(* IEC 61131-3 sources: PLC_I/plc/src/application, 8 files *)

(* ---- 结构体_运行时.st ---- *)
(* Volatile exchange. Call Server before installed axis consumers each scan.
   ConsumerMask proves program routing, never physical online or safety status. *)
TYPE 结构体_运行时 :
STRUCT
    ast轴 : ARRAY[0..15] OF 结构体_轴状态;
    aw轴命令 : ARRAY[0..15] OF WORD;
    aw轴序列 : ARRAY[0..15] OF WORD;
    adi轴目标 : ARRAY[0..15] OF DINT;
    audi轴速度 : ARRAY[0..15] OF UDINT;
    audi轴加速度 : ARRAY[0..15] OF UDINT;
    audi轴减速度 : ARRAY[0..15] OF UDINT;
    audi轴停止减速度 : ARRAY[0..15] OF UDINT;
    w轴消费掩码 : WORD;
    ast气缸 : ARRAY[0..53] OF 结构体_气缸状态;
    aw气缸命令 : ARRAY[0..53] OF WORD;
    aw气缸序列 : ARRAY[0..53] OF WORD;
    b手动 : BOOL;
    b运行 : BOOL;
    b暂停 : BOOL;
    bHMI在线 : BOOL;
    b复位中 : BOOL;
    (* 上位机命令 2/3/4 的一扫描事件。服务端在受理的同一扫描置位，
       PRG 在下一扫描消费后清零；与物理按钮沿分开，避免被 R_TRIG 合并。 *)
    b启动脉冲 : BOOL;
    b暂停脉冲 : BOOL;
    b恢复脉冲 : BOOL;
    b硬急停 : BOOL;
    b软急停 : BOOL;
    b待复位 : BOOL := TRUE;
    ui输入点数 : UINT;
    ui输出点数 : UINT;
    aw输入 : ARRAY[0..7] OF WORD;
    aw输出 : ARRAY[0..7] OF WORD;
END_STRUCT
END_TYPE

(* ---- 全局变量_错误码.gvl.st ---- *)
(* 拒绝/错误码集中定义。FB 只引用名称，避免数字散落各文件。
   数值与协议 register-map 的拒绝码一致，新增码必须同步协议表。 *)
VAR_GLOBAL CONSTANT
    ERR_已受理   : WORD := 0;
    ERR_签名     : WORD := 1;
    ERR_通信离线 : WORD := 2;
    ERR_急停     : WORD := 3;
    ERR_未绑定   : WORD := 4;
    ERR_离线     : WORD := 5;
    ERR_未使能   : WORD := 6;
    ERR_模式     : WORD := 7;
    ERR_复位中   : WORD := 8;
    ERR_参数     : WORD := 9;
    ERR_忙       : WORD := 10;
    ERR_待复位   : WORD := 11;
    ERR_正式流程 : WORD := 12;
    ERR_未接入   : WORD := 14;
    ERR_非法     : WORD := 15;
    ERR_纪元     : WORD := 16;
    ERR_故障     : WORD := 17;
    ERR_无点位   : WORD := 18;
    ERR_取消     : WORD := 19;
    ERR_定标     : WORD := 20;
    ERR_软限位   : WORD := 21;
    ERR_速度     : WORD := 22;
    ERR_P0       : WORD := 26;
    ERR_目标越限 : WORD := 27;
    ERR_速度无效 : WORD := 28;
END_VAR

(* ---- 函数_动作许可.st ---- *)
(* Sole action-permission boundary (SBR_动作许可 role). Structural validation
   belongs to 函数_校验, never duplicate movement predicates in HMI. *)
FUNCTION 函数_动作许可 : WORD
VAR_INPUT
    Code : WORD;
    ObjectWord : WORD;
    HmiOnline : BOOL;
    JogBusy : BOOL;
    Resetting : BOOL;
    b自动请求 : BOOL := FALSE;
    b气缸已受理 : BOOL := FALSE; (* 仅驱动消费时复核当前许可 *)
    b暂停恢复 : BOOL := FALSE; (* 仅暂停恢复FB的轴27，允许在暂停状态回快照 *)
    b恢复已下发 : BOOL := FALSE; (* 持续复核时忽略本动作自身的Busy *)
    di恢复目标 : DINT := 0;
END_VAR
VAR_IN_OUT
    Runtime : 结构体_运行时;
    Store : 结构体_配置;
END_VAR
VAR
    w类别 : WORD;
    ui对象索引 : UINT;
    ui轴号 : UINT;
    w归属 : WORD;
    b空闲槽 : BOOL;
    b对象已绑定 : BOOL;
    b硬件已接入 : BOOL;
    b是停止 : BOOL;
    b有点位 : BOOL;
    i循环 : UINT;
    i子循环 : UINT;
    di正限位 : DINT;
    di负限位 : DINT;
    di位置 : DINT;
    dw值 : DWORD;
END_VAR

函数_动作许可 := ERR_已受理;
w类别 := SHR(ObjectWord, 8);
ui对象索引 := WORD_TO_UINT(ObjectWord AND 16#00FF);
IF (w类别 > 3) OR ((w类别 = 0) AND (ui对象索引 <> 0))
OR ((w类别 = 1) AND (ui对象索引 >= 16))
OR ((w类别 = 2) AND (ui对象索引 >= 54))
OR ((w类别 = 3) AND (ui对象索引 >= 120)) THEN
    函数_动作许可 := ERR_非法; RETURN;
END_IF;
IF b暂停恢复 AND ((w类别 <> 1) OR (Code <> 27)) THEN
    函数_动作许可 := ERR_非法; RETURN;
END_IF;
ui轴号 := ui对象索引;
b空闲槽 := FALSE;
IF w类别 = 3 THEN
    b空闲槽 := Store.aw点位[ui对象索引, 4] = XJV1_POINT_FREE;
    w归属 := SHR(Store.aw点位[ui对象索引, 4], 2) AND WORD#16#000F;
    ui轴号 := WORD_TO_UINT(w归属);
END_IF;
b对象已绑定 := w类别 = 0;
b硬件已接入 := (Runtime.w轴消费掩码 AND w已绑定轴) = w已绑定轴;
IF w类别 = 1 THEN
    b对象已绑定 := (w已绑定轴 AND SHL(WORD#1, ui轴号)) <> 0;
    b硬件已接入 := (Runtime.w轴消费掩码 AND SHL(WORD#1, ui轴号)) <> 0;
ELSIF w类别 = 3 THEN
    (* An owned point is bound exactly when its owner axis is bound; free
       slots are handled separately below. *)
    b对象已绑定 := NOT b空闲槽 AND ((w已绑定轴 AND SHL(WORD#1, ui轴号)) <> 0);
    b硬件已接入 := (Runtime.w轴消费掩码 AND SHL(WORD#1, ui轴号)) <> 0;
ELSIF w类别 = 2 THEN
    b对象已绑定 := (lw已绑定气缸 AND SHL(LWORD#1, ui对象索引)) <> 0;
    b硬件已接入 := ab气缸映射有效[ui对象索引];
END_IF;
b是停止 := (Code = 9) OR (Code = 10) OR (Code = 26) OR (Code = 42);
(* Stop codes bypass every ordinary gate; an unbound object still rejects 4. *)
IF b是停止 THEN
    IF NOT b对象已绑定 THEN 函数_动作许可 := ERR_未绑定; END_IF;
    RETURN;
END_IF;
IF NOT HmiOnline THEN 函数_动作许可 := ERR_通信离线; RETURN; END_IF;
IF (w类别 = 3) AND b空闲槽 THEN
    (* Free pool slot: only a code-50 claim may address it; the candidate
       owner axis is validated against the binding table in Config. *)
    IF Code <> 50 THEN 函数_动作许可 := ERR_未绑定; RETURN; END_IF;
    IF Runtime.b硬急停 OR Runtime.b软急停 THEN 函数_动作许可 := ERR_急停; RETURN; END_IF;
    IF Resetting THEN 函数_动作许可 := ERR_复位中; RETURN; END_IF;
    IF NOT Runtime.b手动 THEN 函数_动作许可 := ERR_模式; RETURN; END_IF;
    RETURN;
END_IF;
IF Code = 53 THEN 函数_动作许可 := ERR_未接入; RETURN; END_IF;
IF Code = 11 THEN
    (* Clear only the software latch. This does not grant motion permission,
       reset faults, enable an axis, or resume the sequence. *)
    IF Runtime.b硬急停 THEN 函数_动作许可 := ERR_急停; END_IF;
    RETURN;
END_IF;
IF Runtime.b硬急停 OR Runtime.b软急停 THEN 函数_动作许可 := ERR_急停; RETURN; END_IF;
IF NOT b对象已绑定 THEN 函数_动作许可 := ERR_未绑定; RETURN; END_IF;
IF w类别 = 2 THEN
    IF Resetting THEN 函数_动作许可 := ERR_复位中; RETURN; END_IF;
    IF Runtime.b暂停 THEN 函数_动作许可 := ERR_模式; RETURN; END_IF;
    IF b自动请求 THEN
        IF NOT 全局变量_运行配置.b正式流程已接入 THEN 函数_动作许可 := ERR_正式流程; RETURN; END_IF;
        IF NOT Runtime.b运行 THEN 函数_动作许可 := ERR_模式; RETURN; END_IF;
    ELSIF NOT Runtime.b手动 THEN 函数_动作许可 := ERR_模式; RETURN;
    END_IF;
    IF (Code <> 40) AND (Code <> 41) AND (Code <> 50) THEN 函数_动作许可 := ERR_未接入; RETURN; END_IF;
    IF NOT b气缸已受理 AND (全局变量_气缸请求.ast请求[ui对象索引].b忙
        OR Runtime.ast气缸[ui对象索引].b运动中) THEN 函数_动作许可 := ERR_忙; RETURN; END_IF;
    IF Code = 50 THEN RETURN; END_IF;
    IF NOT b硬件已接入 THEN 函数_动作许可 := ERR_未接入; RETURN; END_IF;
    IF NOT ab气缸模块就绪[ui对象索引] THEN 函数_动作许可 := ERR_离线; RETURN; END_IF;
    IF Runtime.ast气缸[ui对象索引].b故障 THEN 函数_动作许可 := ERR_故障; RETURN; END_IF;
    (* 手动调试不依赖上电复位和现场配置确认：手动模式下可以直接触发
       动点/原点。自动请求仍必须完成确认与复位，避免工艺在未确认配置上运行。 *)
    IF b自动请求 THEN
        IF Runtime.b待复位 THEN 函数_动作许可 := ERR_待复位; RETURN; END_IF;
        IF NOT Store.b已确认 THEN 函数_动作许可 := ERR_未接入; RETURN; END_IF;
    END_IF;
    IF NOT 气缸_配置有效(缸号 := ui对象索引, Store := Store) THEN 函数_动作许可 := ERR_参数; END_IF;
    RETURN;
END_IF;
(* 整机启动/暂停/恢复。正式工艺未接入时三条一律拒绝 12，与原程序
   “NOT b正式流程已接入 → 拒绝” 一致；接入后由运行状态机判定模式与暂停，
   这里只做安全与前置条件检查，不复制运行状态机的优先级逻辑。 *)
IF (Code = 2) OR (Code = 3) OR (Code = 4) THEN
    IF NOT 全局变量_运行配置.b正式流程已接入 THEN 函数_动作许可 := ERR_正式流程; RETURN; END_IF;
    IF Code = 2 THEN
        IF Runtime.b待复位 THEN 函数_动作许可 := ERR_未接入; RETURN; END_IF;
    ELSIF Code = 4 THEN
        IF NOT Runtime.b暂停 THEN 函数_动作许可 := ERR_未接入; RETURN; END_IF;
    END_IF;
    RETURN;
END_IF;
IF Resetting AND (Code <> 21) THEN 函数_动作许可 := ERR_复位中; RETURN; END_IF;
IF w类别 = 0 THEN
    IF Code = 1 THEN
        IF NOT b硬件已接入 THEN 函数_动作许可 := ERR_未接入; RETURN; END_IF;
        FOR i循环 := 0 TO 15 DO
            IF (w已绑定轴 AND SHL(WORD#1, i循环)) <> 0 THEN
                IF NOT Runtime.ast轴[i循环].b在线 THEN 函数_动作许可 := ERR_离线; RETURN; END_IF;
            END_IF;
        END_FOR;
    ELSIF Code = 52 THEN
        IF NOT Runtime.b手动 THEN 函数_动作许可 := ERR_模式; RETURN; END_IF;
        FOR i循环 := 0 TO 15 DO
            IF (w已绑定轴 AND SHL(WORD#1, i循环)) <> 0 THEN
                IF NOT Runtime.ast轴[i循环].b在线 THEN 函数_动作许可 := ERR_离线; RETURN; END_IF;
                IF Runtime.ast轴[i循环].b故障 THEN 函数_动作许可 := ERR_故障; RETURN; END_IF;
                IF Runtime.ast轴[i循环].b运动中 OR NOT Runtime.ast轴[i循环].b静止 THEN
                    函数_动作许可 := ERR_忙; RETURN;
                END_IF;
                di正限位 := DWORD_TO_DINT(SHL(WORD_TO_DWORD(Store.aw轴配置[i循环, 0]), 16) OR WORD_TO_DWORD(Store.aw轴配置[i循环, 1]));
                di负限位 := DWORD_TO_DINT(SHL(WORD_TO_DWORD(Store.aw轴配置[i循环, 2]), 16) OR WORD_TO_DWORD(Store.aw轴配置[i循环, 3]));
                IF (Store.aw轴配置[i循环, 14] <> 1) OR (Store.aw轴配置[i循环, 15] <> 0) THEN
                    函数_动作许可 := ERR_定标; RETURN;
                END_IF;
                IF di负限位 >= di正限位 THEN 函数_动作许可 := ERR_软限位; RETURN; END_IF;
                FOR i子循环 := 2 TO 6 DO
                    dw值 := SHL(WORD_TO_DWORD(Store.aw轴配置[i循环, i子循环 * 2]), 16) OR WORD_TO_DWORD(Store.aw轴配置[i循环, i子循环 * 2 + 1]);
                    IF (dw值 = 0) OR (dw值 > DWORD#2147483647) THEN
                        函数_动作许可 := 函数_参数码(i子循环); RETURN;
                    END_IF;
                    IF NOT 函数_额定值(AxisIndex := i循环, Field := i子循环,
                        Value := DWORD_TO_UDINT(dw值)) THEN
                        函数_动作许可 := 函数_参数码(i子循环); RETURN;
                    END_IF;
                END_FOR;
                (* Standby point P0 of axis i is pool slot i by definition. *)
                IF (SHR(Store.aw点位[i循环, 4], 2) AND WORD#16#000F) <> UINT_TO_WORD(i循环)
                OR (Store.aw点位[i循环, 4] AND 3) <> 3 THEN 函数_动作许可 := ERR_无点位; RETURN; END_IF;
                di位置 := DWORD_TO_DINT(SHL(WORD_TO_DWORD(Store.aw点位[i循环, 0]), 16) OR WORD_TO_DWORD(Store.aw点位[i循环, 1]));
                dw值 := SHL(WORD_TO_DWORD(Store.aw点位[i循环, 2]), 16) OR WORD_TO_DWORD(Store.aw点位[i循环, 3]);
                IF (di位置 < di负限位) OR (di位置 > di正限位) THEN 函数_动作许可 := ERR_P0; RETURN; END_IF;
                IF (dw值 = 0) OR (dw值 > DWORD#2147483647) THEN 函数_动作许可 := ERR_速度无效; RETURN; END_IF;
            END_IF;
        END_FOR;
        FOR i循环 := 0 TO 53 DO
            IF (lw已绑定气缸 AND SHL(LWORD#1, i循环)) <> 0 THEN
                IF NOT 气缸_配置有效(缸号 := i循环, Store := Store) THEN 函数_动作许可 := ERR_参数; RETURN; END_IF;
                IF 全局变量_气缸请求.ast请求[i循环].b忙 THEN 函数_动作许可 := ERR_忙; RETURN; END_IF;
            END_IF;
        END_FOR;
    ELSE
        函数_动作许可 := ERR_未接入;
    END_IF;
    RETURN;
END_IF;
IF (Runtime.aw轴命令[ui轴号] <> 0) AND (Code <> 21) THEN
    函数_动作许可 := ERR_忙; RETURN;
END_IF;
IF NOT b自动请求 AND 全局变量_轴请求.ast请求[ui轴号].b忙 AND (Code <> 21) THEN
    函数_动作许可 := ERR_忙; RETURN;
END_IF;
CASE Code OF
    20, 21, 22, 23, 24, 25, 27, 28, 29, 30, 31, 50: ;
ELSE
    函数_动作许可 := ERR_未接入; RETURN;
END_CASE;
IF NOT Runtime.ast轴[ui轴号].b在线 THEN 函数_动作许可 := ERR_离线; RETURN; END_IF;
(* 硬限位未接线时必须保留软限位，否则拒绝运动类命令，避免无边界保护。 *)
IF (Code = 22) OR (Code = 24) OR (Code = 25) OR (Code = 27)
    OR (Code = 28) OR (Code = 29) THEN
    IF NOT 全局变量_运行配置.b硬限位已接线
        AND ((Store.aw轴配置[ui轴号, 14] AND WORD#16#0001) = 0) THEN
        函数_动作许可 := ERR_未接入; RETURN;
    END_IF;
END_IF;
(* 写参数（31/50）不动轴，报警期间也允许改；复位 23 与去使能 21 同样放行。 *)
IF Runtime.ast轴[ui轴号].b故障 AND (Code <> 21) AND (Code <> 23)
    AND (Code <> 31) AND (Code <> 50) THEN
    函数_动作许可 := ERR_故障; RETURN;
END_IF;
IF b暂停恢复 THEN
    (* 恢复有独立模式条件；不能借普通自动许可放开暂停中的其他命令。 *)
    IF NOT 全局变量_运行配置.b正式流程已接入 THEN 函数_动作许可 := ERR_正式流程; RETURN; END_IF;
    (* 运行控制在暂停时发布手动模式，恢复仍以暂停握手为准。 *)
    IF NOT Runtime.b暂停 THEN 函数_动作许可 := ERR_模式; RETURN; END_IF;
    IF Runtime.b待复位 THEN 函数_动作许可 := ERR_待复位; RETURN; END_IF;
    di正限位 := DWORD_TO_DINT(SHL(WORD_TO_DWORD(Store.aw轴配置[ui轴号, 0]), 16) OR WORD_TO_DWORD(Store.aw轴配置[ui轴号, 1]));
    di负限位 := DWORD_TO_DINT(SHL(WORD_TO_DWORD(Store.aw轴配置[ui轴号, 2]), 16) OR WORD_TO_DWORD(Store.aw轴配置[ui轴号, 3]));
    IF (Store.aw轴配置[ui轴号, 14] AND 1) <> 0 THEN
        IF (di负限位 >= di正限位) OR (di恢复目标 < di负限位) OR (di恢复目标 > di正限位) THEN
            函数_动作许可 := ERR_软限位; RETURN;
        END_IF;
    END_IF;
    IF ((di恢复目标 > Runtime.ast轴[ui轴号].di位置) AND ((Runtime.ast轴[ui轴号].w限位 AND 5) <> 0))
        OR ((di恢复目标 < Runtime.ast轴[ui轴号].di位置) AND ((Runtime.ast轴[ui轴号].w限位 AND 10) <> 0)) THEN
        函数_动作许可 := ERR_故障; RETURN;
    END_IF;
ELSIF b自动请求 THEN
    IF NOT 全局变量_运行配置.b正式流程已接入 THEN 函数_动作许可 := ERR_正式流程; RETURN; END_IF;
    IF NOT Runtime.b运行 OR Runtime.b暂停 THEN 函数_动作许可 := ERR_模式; RETURN; END_IF;
    IF Runtime.b待复位 THEN 函数_动作许可 := ERR_待复位; RETURN; END_IF;
ELSIF NOT Runtime.b手动 AND (Code <> 21) THEN 函数_动作许可 := ERR_模式; RETURN;
END_IF;
IF ((Code = 22) OR (Code = 24) OR (Code = 25) OR (Code = 27) OR (Code = 28) OR (Code = 29) OR (Code = 30))
AND NOT Runtime.ast轴[ui轴号].b已使能 THEN 函数_动作许可 := ERR_未使能; RETURN; END_IF;
(* 清故障在报警态必须可重试：轴停在 ErrorStop 时 b运动中 可能因残留停止阶段为真，
   若因此拒绝 23，现场就永远清不掉。复位本身仍要求 MC_Reset 成功。 *)
IF (Code >= 20) AND (Code <= 30) AND (Code <> 21)
AND NOT (b暂停恢复 AND b恢复已下发)
AND NOT Runtime.ast轴[ui轴号].b可下发 THEN
    函数_动作许可 := ERR_忙; RETURN;
END_IF;
IF (Runtime.ast轴[ui轴号].b运动中 OR NOT Runtime.ast轴[ui轴号].b静止) AND (Code <> 21) AND (Code <> 23)
    AND NOT (b暂停恢复 AND b恢复已下发) THEN
    函数_动作许可 := ERR_忙; RETURN;
END_IF;
IF (Code = 24) OR (Code = 25) THEN
    IF JogBusy THEN 函数_动作许可 := ERR_忙; RETURN; END_IF;
    IF ((Code = 24) AND ((Runtime.ast轴[ui轴号].w限位 AND 5) <> 0))
    OR ((Code = 25) AND ((Runtime.ast轴[ui轴号].w限位 AND 10) <> 0)) THEN
        函数_动作许可 := ERR_故障; RETURN;
    END_IF;
END_IF;
IF Code = 29 THEN
    b有点位 := FALSE;
    FOR i循环 := 0 TO 119 DO
        b有点位 := b有点位 OR ((SHR(Store.aw点位[i循环, 4], 2) AND WORD#16#000F) = UINT_TO_WORD(ui轴号)
            AND ((Store.aw点位[i循环, 4] AND 3) = 3));
    END_FOR;
    IF NOT b有点位 THEN 函数_动作许可 := ERR_无点位; RETURN; END_IF;
END_IF;
IF ((Code >= 20) AND (Code <= 30)) AND NOT b硬件已接入 THEN
    函数_动作许可 := ERR_未接入; RETURN;
END_IF;
IF (Code = 20) OR (Code = 22) OR (Code = 24) OR (Code = 25)
OR (Code = 27) OR (Code = 28) OR (Code = 29) THEN
    FOR i子循环 := 2 TO 6 DO
        dw值 := SHL(WORD_TO_DWORD(Store.aw轴配置[ui轴号, i子循环 * 2]), 16)
            OR WORD_TO_DWORD(Store.aw轴配置[ui轴号, i子循环 * 2 + 1]);
        IF NOT 函数_额定值(AxisIndex := ui轴号, Field := i子循环,
            Value := DWORD_TO_UDINT(dw值)) THEN
            函数_动作许可 := 函数_参数码(i子循环); RETURN;
        END_IF;
    END_FOR;
END_IF;
END_FUNCTION

(* ---- 功能块_暂停恢复.st ---- *)
(* 暂停快照与恢复。移植自原程序“暂停快照 / 暂停回位”三段，只保留必要行为：

   暂停沿 -> 对运动中轴下受控停止 26 -> 全部静止后抓拍位置
   恢复请求 -> 对偏离超过容差的轴下发绝对定位 27 回快照位置 -> 结果 2 即完成
   急停 / 轴离线或故障 -> 立即判失败并撤销本块下发的命令

   不产生动作许可，不替代 功能块_轴 的安全判定。
   必须在 功能块_服务端 之后、各轴消费之前调用（服务端每扫描开头清零命令数组）。 *)
FUNCTION_BLOCK 功能块_暂停恢复
VAR_INPUT
    b暂停 : BOOL;
    b请求 : BOOL;
    b急停 : BOOL;
    di容差 : DINT;
    (* 停稳确认时间。原程序为 300 ms；做成输入便于自测用更短的值，
       现场调用保持 300 ms。 *)
    di停稳ms : DINT;
END_VAR
VAR_IN_OUT
    Runtime : 结构体_运行时;
END_VAR
VAR_OUTPUT
    b恢复中 : BOOL;
    b恢复完成 : BOOL;
    b恢复失败 : BOOL;
    b曾偏离 : BOOL;
    b已抓拍 : BOOL;
    (* 内部阶段只读发布，供上位机诊断与自测观察。 *)
    ui内部阶段 : UINT;
END_VAR
VAR
    i阶段 : UINT; (* 0 空闲，1 停车等待静止，2 已抓拍待恢复，3 回位中 *)
    b暂停上周期 : BOOL;
    b请求上周期 : BOOL;
    b请求沿 : BOOL;
    adi快照 : ARRAY[0..15] OF DINT;
    (* 只有收到本轮回位 27 的轴才参与完成判定；未偏离的轴不动作，
       不能被当成“未到位”而把恢复永久卡住。 *)
    ab已下发 : ARRAY[0..15] OF BOOL;
    w序列 : WORD;
    b暂停沿 : BOOL;
    b封锁 : BOOL;
    b全部静止 : BOOL;
    b全部到位 : BOOL;
    b取消恢复 : BOOL;
    b恢复动作存在 : BOOL;
    w许可 : WORD;
    tmr停稳 : TON;
    tmr恢复 : TON;
    i循环 : UINT;
END_VAR

b恢复中 := FALSE;
b取消恢复 := (i阶段 = 3) AND (NOT b暂停 OR NOT b请求);
(* b已抓拍 是锁存状态，不是脉冲：暂停沿/解除时清零，抓拍成功时置位。
   上位机与自测都靠它判断“快照是否有效”，脉冲化会漏读。 *)
b暂停沿 := b暂停 AND NOT b暂停上周期;
b暂停上周期 := b暂停;
b请求沿 := b请求 AND NOT b请求上周期;
b请求上周期 := b请求;

(* 安全条件不满足时任何恢复都不成立。 *)
b封锁 := b急停 OR Runtime.b硬急停 OR Runtime.b软急停;
IF b请求沿 OR (i阶段 = 3) THEN
    b封锁 := b封锁 OR NOT Runtime.bHMI在线 OR Runtime.b待复位 OR Runtime.b复位中
        OR NOT 全局变量_运行配置.b正式流程已接入;
END_IF;
FOR i循环 := 0 TO 15 DO
    IF (w已绑定轴 AND SHL(WORD#1, i循环)) <> 0 THEN
        b封锁 := b封锁 OR NOT Runtime.ast轴[i循环].b在线 OR Runtime.ast轴[i循环].b故障;
    END_IF;
END_FOR;
(* 先完整预检全部目标，再发任何轴；回位中每扫描继续复核。
   使用LINT比较，DINT极值两端相减不会溢出。 *)
IF ((i阶段 = 2) AND b请求沿) OR (i阶段 = 3) THEN
    FOR i循环 := 0 TO 15 DO
        IF (w已绑定轴 AND SHL(WORD#1, i循环)) <> 0 THEN
            IF ab已下发[i循环] OR
                (ABS(DINT_TO_LINT(Runtime.ast轴[i循环].di位置) - DINT_TO_LINT(adi快照[i循环])) > DINT_TO_LINT(di容差)) THEN
                w许可 := 函数_动作许可(Code := 27, ObjectWord := WORD#16#0100 OR UINT_TO_WORD(i循环),
                    HmiOnline := Runtime.bHMI在线, JogBusy := FALSE, Resetting := Runtime.b复位中,
                    b暂停恢复 := TRUE, b恢复已下发 := (i阶段 = 3) AND ab已下发[i循环],
                    di恢复目标 := adi快照[i循环], Runtime := Runtime, Store := 全局变量_保持区.Store);
                b封锁 := b封锁 OR (w许可 <> 0);
            END_IF;
        END_IF;
    END_FOR;
END_IF;
IF (i阶段 = 3) AND b封锁 THEN b取消恢复 := TRUE; END_IF;

IF b暂停沿 THEN
    i阶段 := 1;
    b曾偏离 := FALSE;
    b恢复完成 := FALSE;
    b恢复失败 := FALSE;
    b已抓拍 := FALSE;
    w序列 := w序列 + 1;
    tmr停稳(IN := FALSE, PT := DINT_TO_TIME(di停稳ms));
    FOR i循环 := 0 TO 15 DO
        adi快照[i循环] := Runtime.ast轴[i循环].di位置;
        ab已下发[i循环] := FALSE;
    END_FOR;
ELSIF NOT b暂停 THEN
    i阶段 := 0;
    b曾偏离 := FALSE;
    b已抓拍 := FALSE;
END_IF;

CASE i阶段 OF
    1:
        (* 受控停止。序列固定，重复下发同一序列不会在轴内重复触发。 *)
        b全部静止 := TRUE;
        FOR i循环 := 0 TO 15 DO
            IF (w已绑定轴 AND SHL(WORD#1, i循环)) <> 0 THEN
                IF Runtime.ast轴[i循环].b运动中 OR NOT Runtime.ast轴[i循环].b静止 THEN
                    b全部静止 := FALSE;
                    Runtime.aw轴命令[i循环] := 26;
                    Runtime.aw轴序列[i循环] := w序列;
                END_IF;
            END_IF;
        END_FOR;
        tmr停稳(IN := b全部静止 AND NOT b封锁, PT := DINT_TO_TIME(di停稳ms));
        IF tmr停稳.Q THEN
            (* 停稳后重新抓拍：减速距离不算偏离。 *)
            FOR i循环 := 0 TO 15 DO adi快照[i循环] := Runtime.ast轴[i循环].di位置; END_FOR;
            b已抓拍 := TRUE;
            i阶段 := 2;
        END_IF;
    2:
        (* 暂停期间只监视偏离，不自动动作。 *)
        FOR i循环 := 0 TO 15 DO
            IF (w已绑定轴 AND SHL(WORD#1, i循环)) <> 0 THEN
                IF ABS(DINT_TO_LINT(Runtime.ast轴[i循环].di位置) - DINT_TO_LINT(adi快照[i循环])) > DINT_TO_LINT(di容差) THEN
                    b曾偏离 := TRUE;
                END_IF;
            END_IF;
        END_FOR;
        (* 恢复请求只在上升沿处理一次：b请求 是电平，重复处理会每扫描
           重新下发 27，命令槽无法释放，安全封锁时也撤不干净。 *)
        IF b请求沿 AND b封锁 THEN b恢复失败 := TRUE; END_IF;
        IF b请求沿 AND NOT b封锁 THEN
            b恢复完成 := FALSE;
            b恢复失败 := FALSE;
            b恢复动作存在 := FALSE;
            FOR i循环 := 0 TO 15 DO
                IF ((w已绑定轴 AND SHL(WORD#1, i循环)) <> 0)
                    AND (ABS(DINT_TO_LINT(Runtime.ast轴[i循环].di位置) - DINT_TO_LINT(adi快照[i循环])) > DINT_TO_LINT(di容差)) THEN
                    b恢复动作存在 := TRUE;
                END_IF;
            END_FOR;
            IF b恢复动作存在 THEN
                w序列 := w序列 + 1;
                FOR i循环 := 0 TO 15 DO ab已下发[i循环] := FALSE; END_FOR;
                FOR i循环 := 0 TO 15 DO
                    IF (w已绑定轴 AND SHL(WORD#1, i循环)) <> 0 THEN
                        IF ABS(DINT_TO_LINT(Runtime.ast轴[i循环].di位置) - DINT_TO_LINT(adi快照[i循环])) > DINT_TO_LINT(di容差) THEN
                            (* 回位参数取保持配置，与命令 27 的下发参数同源。 *)
                            Runtime.adi轴目标[i循环] := adi快照[i循环];
                            Runtime.audi轴速度[i循环] := DWORD_TO_UDINT(
                                SHL(WORD_TO_DWORD(全局变量_保持区.Store.aw轴配置[i循环, 4]), 16)
                                OR WORD_TO_DWORD(全局变量_保持区.Store.aw轴配置[i循环, 5]));
                            Runtime.audi轴加速度[i循环] := DWORD_TO_UDINT(
                                SHL(WORD_TO_DWORD(全局变量_保持区.Store.aw轴配置[i循环, 8]), 16)
                                OR WORD_TO_DWORD(全局变量_保持区.Store.aw轴配置[i循环, 9]));
                            Runtime.audi轴减速度[i循环] := DWORD_TO_UDINT(
                                SHL(WORD_TO_DWORD(全局变量_保持区.Store.aw轴配置[i循环, 10]), 16)
                                OR WORD_TO_DWORD(全局变量_保持区.Store.aw轴配置[i循环, 11]));
                            Runtime.audi轴停止减速度[i循环] := DWORD_TO_UDINT(
                                SHL(WORD_TO_DWORD(全局变量_保持区.Store.aw轴配置[i循环, 12]), 16)
                                OR WORD_TO_DWORD(全局变量_保持区.Store.aw轴配置[i循环, 13]));
                            Runtime.aw轴命令[i循环] := 27;
                            Runtime.aw轴序列[i循环] := w序列;
                            ab已下发[i循环] := TRUE;
                        END_IF;
                    END_IF;
                END_FOR;
                tmr恢复(IN := FALSE, PT := T#120s);
                i阶段 := 3;
            ELSE
                (* 没偏离就没有要回的位置，恢复直接成立。 *)
                b恢复完成 := TRUE;
            END_IF;
        END_IF;

    3:
        b恢复中 := TRUE;
        b全部到位 := TRUE;
        FOR i循环 := 0 TO 15 DO
            IF (w已绑定轴 AND SHL(WORD#1, i循环)) <> 0 AND ab已下发[i循环] THEN
                b全部到位 := b全部到位 AND (Runtime.ast轴[i循环].w序列 = w序列)
                    AND (Runtime.ast轴[i循环].w运动结果 = 2)
                    AND Runtime.ast轴[i循环].b静止;
            END_IF;
        END_FOR;
        tmr恢复(IN := TRUE, PT := T#120s);
        IF b取消恢复 OR b封锁 OR tmr恢复.Q THEN
            b取消恢复 := TRUE;
            b恢复失败 := TRUE;
            b恢复中 := FALSE;
            i阶段 := 2;
        ELSIF b全部到位 THEN
            FOR i循环 := 0 TO 15 DO ab已下发[i循环] := FALSE; END_FOR;
            b恢复完成 := TRUE;
            b恢复中 := FALSE;
            i阶段 := 2;
        END_IF;
END_CASE;
(* 清命令槽不能取消轴内已锁存的27；主动发26并使用新序列。 *)
IF b取消恢复 THEN
    w序列 := w序列 + 1;
    FOR i循环 := 0 TO 15 DO
        IF ab已下发[i循环] THEN
            Runtime.aw轴命令[i循环] := 26;
            Runtime.aw轴序列[i循环] := w序列;
            ab已下发[i循环] := FALSE;
        END_IF;
    END_FOR;
    b恢复中 := FALSE;
    b恢复完成 := FALSE;
    b恢复失败 := TRUE;
END_IF;
ui内部阶段 := i阶段;
END_FUNCTION_BLOCK

(* ---- 功能块_模式管理.st ---- *)
(* 模式/暂停恢复的唯一状态拥有者。服务端之后、轴组之前调用一次。 *)
FUNCTION_BLOCK 功能块_模式管理
VAR_INPUT StartButton : BOOL; PauseButton : BOOL; ResetButton : BOOL; END_VAR
VAR_IN_OUT Runtime : 结构体_运行时; END_VAR
VAR
    fb运行 : 功能块_运行控制;
    fb暂停恢复 : 功能块_暂停恢复;
    fb启动滤波 : 功能块_输入滤波;
    fb暂停滤波 : 功能块_输入滤波;
    fb复位滤波 : 功能块_输入滤波;
    b复位事件 : BOOL;
    b复位上周期 : BOOL;
    b设备报警 : BOOL;
    b急停 : BOOL;
    i循环 : UINT;
END_VAR
fb启动滤波(b信号 := StartButton, i模式 := 1,
    di滤波时间真 := 全局变量_运行配置.di输入滤波时间ms,
    di滤波时间假 := 全局变量_运行配置.di输入滤波时间ms);
fb暂停滤波(b信号 := PauseButton, i模式 := 1,
    di滤波时间真 := 全局变量_运行配置.di输入滤波时间ms,
    di滤波时间假 := 全局变量_运行配置.di输入滤波时间ms);
fb复位滤波(b信号 := ResetButton, i模式 := 1,
    di滤波时间真 := 全局变量_运行配置.di输入滤波时间ms,
    di滤波时间假 := 全局变量_运行配置.di输入滤波时间ms);
b复位事件 := fb复位滤波.b滤波信号 AND NOT b复位上周期;
b复位上周期 := fb复位滤波.b滤波信号;
b急停 := Runtime.b硬急停;
(* ===== 区域 3：运行模式与命令脉冲消费 ===== *)
(* 运行状态机：物理按钮 + 上位机命令 2/3/4。命令 2 在
   b正式流程已接入 = FALSE 时仍由 函数_动作许可 拒绝为 12。 *)
b设备报警 := FALSE;
FOR i循环 := 0 TO 15 DO
    IF (w已绑定轴 AND SHL(WORD#1, i循环)) <> 0 THEN b设备报警 := b设备报警 OR Runtime.ast轴[i循环].b故障; END_IF;
END_FOR;
fb运行(b初始化完成 := TRUE,
    b系统复位完成 := NOT Runtime.b待复位,
    b系统复位中 := FALSE,
    b系统复位失败 := FALSE,
    b启动按钮 := fb启动滤波.b滤波信号 AND 全局变量_运行配置.b正式流程已接入,
    b暂停按钮 := fb暂停滤波.b滤波信号,
    b启动事件 := Runtime.b启动脉冲,
    b暂停事件 := Runtime.b暂停脉冲,
    (* 物理复位按钮与命令 4 等效：原程序“暂停中按复位进入暂停恢复”。 *)
    b恢复事件 := Runtime.b恢复脉冲 OR (b复位事件 AND 全局变量_运行配置.b正式流程已接入),
    b致命报警 := Runtime.b硬急停 OR Runtime.b软急停 OR b设备报警,
    b急停 := b急停 OR Runtime.b软急停,
    b暂停报警 := b设备报警,
    b预警 := FALSE,
    b暂停恢复中 := fb暂停恢复.b恢复中,
    b暂停恢复完成 := fb暂停恢复.b恢复完成,
    b暂停恢复失败 := fb暂停恢复.b恢复失败,
    b流程完成 := FALSE);
Runtime.b运行 := fb运行.b运行指令;
Runtime.b暂停 := fb运行.b暂停中;
Runtime.b手动 := fb运行.b手动模式;
(* 命令 2/3/4 是一扫描事件：服务端本扫描置位，这里消费后立即清零，
   下一扫描不会重复触发。 *)
Runtime.b启动脉冲 := FALSE;
Runtime.b暂停脉冲 := FALSE;
Runtime.b恢复脉冲 := FALSE;

(* 暂停编排：必须在服务端之后，服务端每扫描开头清零命令数组。 *)
fb暂停恢复(b暂停 := fb运行.b暂停中, b请求 := fb运行.b暂停恢复请求,
    b急停 := b急停,
    di容差 := 全局变量_运行配置.di暂停恢复容差,
    di停稳ms := 全局变量_运行配置.di暂停停稳ms, Runtime := Runtime);

(* Cancel automatic requests before consumers when mode changes in this scan.
   Preserve existing stop/disable/reset pulses from the Server. *)
FOR i循环 := 0 TO 15 DO
    IF 全局变量_轴请求.ast请求[i循环].b忙
    AND 全局变量_轴请求.ast请求[i循环].b已下发
    AND (全局变量_轴请求.ast请求[i循环].w命令 <> 26)
    AND (NOT Runtime.b运行 OR Runtime.b暂停 OR NOT Runtime.bHMI在线
        OR Runtime.b硬急停 OR Runtime.b软急停
        OR Runtime.b待复位 OR Runtime.b复位中) THEN
        IF (Runtime.aw轴命令[i循环] = 0) OR (Runtime.aw轴命令[i循环] = 22)
        OR (Runtime.aw轴命令[i循环] = 27) THEN
            Runtime.aw轴命令[i循环] := 26;
        END_IF;
    END_IF;
END_FOR;

END_FUNCTION_BLOCK

(* ---- 功能块_系统复位.st ---- *)
(* Owns reset phase, committed sequence and timeout. Operation 0 advances once
   before arbitration; 1 accepts reset; 2 cancels immediately during arbitration.
   Start/cancel never advance the timer or phase machine a second time. *)
FUNCTION_BLOCK 功能块_系统复位
VAR_INPUT
    Operation : UINT;
    Sequence : WORD;
END_VAR
VAR_IN_OUT
    Runtime : 结构体_运行时;
END_VAR
VAR_OUTPUT
    Busy : BOOL;
    StopRequested : BOOL;
    Failed : BOOL;
END_VAR
VAR
    ui复位阶段 : UINT;
    w复位序列 : WORD;
    b复位完成 : BOOL;
    b复位失败 : BOOL;
    tmr复位 : TON;
    i循环 : UINT;
END_VAR

StopRequested := FALSE;
Failed := FALSE;
CASE Operation OF
    1:
        Runtime.b待复位 := TRUE;
        w复位序列 := Sequence;
        ui复位阶段 := 1;
        StopRequested := TRUE;
    2:
        ui复位阶段 := 0;
    0:
        tmr复位(IN := ui复位阶段 <> 0, PT := T#30s);
        b复位失败 := Runtime.b硬急停 OR Runtime.b软急停 OR tmr复位.Q;
        FOR i循环 := 0 TO 15 DO
            IF (w已绑定轴 AND SHL(WORD#1, i循环)) <> 0 THEN
                b复位失败 := b复位失败 OR NOT Runtime.ast轴[i循环].b在线;
            END_IF;
        END_FOR;
        IF (ui复位阶段 <> 0) AND b复位失败 THEN
            ui复位阶段 := 0;
            Runtime.b待复位 := TRUE;
            StopRequested := TRUE;
            Failed := TRUE;
        END_IF;
        CASE ui复位阶段 OF
            1:
                b复位完成 := TRUE;
                FOR i循环 := 0 TO 15 DO
                    IF (w已绑定轴 AND SHL(WORD#1, i循环)) <> 0 THEN
                        b复位完成 := b复位完成 AND NOT Runtime.ast轴[i循环].b运动中
                            AND Runtime.ast轴[i循环].b可下发
                            AND (Runtime.ast轴[i循环].b静止 OR (Runtime.ast轴[i循环].b故障 AND (Runtime.ast轴[i循环].di速度 = 0)));
                    END_IF;
                END_FOR;
                IF b复位完成 THEN ui复位阶段 := 2; END_IF;
            2:
                FOR i循环 := 0 TO 15 DO
                    IF (w已绑定轴 AND SHL(WORD#1, i循环)) <> 0 THEN
                        Runtime.aw轴命令[i循环] := 23;
                        Runtime.aw轴序列[i循环] := w复位序列;
                    END_IF;
                END_FOR;
                ui复位阶段 := 3;
            3:
                b复位完成 := TRUE;
                FOR i循环 := 0 TO 15 DO
                    IF (w已绑定轴 AND SHL(WORD#1, i循环)) <> 0 THEN
                        b复位完成 := b复位完成 AND (Runtime.ast轴[i循环].w序列 = w复位序列)
                            AND (Runtime.ast轴[i循环].w运动结果 = 2) AND NOT Runtime.ast轴[i循环].b故障
                            AND Runtime.ast轴[i循环].b静止 AND NOT Runtime.ast轴[i循环].b运动中;
                    END_IF;
                END_FOR;
                IF b复位完成 THEN Runtime.b待复位 := FALSE; ui复位阶段 := 4; END_IF;
            4: ui复位阶段 := 0;
        END_CASE;
END_CASE;
Busy := ui复位阶段 <> 0;
END_FUNCTION_BLOCK

(* ---- 功能块_输入滤波.st ---- *)
(* 现场输入去抖。语义与原程序 功能块_输入滤波 一致：
   模式 0 直通；模式 1 按真/假时间分别计时，先到者生效。
   安全输入（急停 X3）不经过本块，避免滤波延迟安全响应。
   X0/X1/X2 走 20 ms 去抖，与原程序 子程序_IO映射__采集 一致。 *)
FUNCTION_BLOCK 功能块_输入滤波
VAR_INPUT
    b信号 : BOOL;
    i模式 : INT; (* 0 = 直通，1 = 去抖 *)
    di滤波时间真 : DINT; (* ms *)
    di滤波时间假 : DINT; (* ms *)
END_VAR
VAR_OUTPUT
    b滤波信号 : BOOL;
END_VAR
VAR
    tmr延时真 : TON;
    tmr延时假 : TON;
END_VAR

CASE i模式 OF
    0:
        tmr延时真(IN := FALSE, PT := DINT_TO_TIME(di滤波时间真));
        tmr延时假(IN := FALSE, PT := DINT_TO_TIME(di滤波时间假));
        b滤波信号 := b信号;
    1:
        tmr延时真(IN := b信号, PT := DINT_TO_TIME(di滤波时间真));
        tmr延时假(IN := NOT b信号, PT := DINT_TO_TIME(di滤波时间假));

        IF tmr延时真.Q THEN
            b滤波信号 := TRUE;
        END_IF;

        IF tmr延时假.Q THEN
            b滤波信号 := FALSE;
        END_IF;
ELSE
    (* 非法模式按直通处理，绝不因为配置错误把一个输入永久锁死。 *)
    tmr延时真(IN := FALSE, PT := DINT_TO_TIME(di滤波时间真));
    tmr延时假(IN := FALSE, PT := DINT_TO_TIME(di滤波时间假));
    b滤波信号 := b信号;
END_CASE;
END_FUNCTION_BLOCK

(* ---- 功能块_运行控制.st ---- *)
(* 整机运行状态机。移植自原程序 功能块_运行控制 + 子程序_运行管理__暂停恢复
   的进入/退出部分，语义逐条对齐：
   优先级 硬故障 > 流程完成 > 初始化/复位 > 暂停 > 启动；
   同一扫描启动与暂停同时出现时暂停优先；
   自动启动必须先通过 b自动可运行（初始化、复位完成、无致命报警、无暂停恢复中）。
   本块只产生“模式与运行指令”，不产生任何动作许可；动作许可仍由
   函数_动作许可 单层判定。 *)
FUNCTION_BLOCK 功能块_运行控制
VAR_INPUT
    b初始化完成 : BOOL;
    b系统复位完成 : BOOL;
    b系统复位中 : BOOL;
    b系统复位失败 : BOOL;
    (* 物理按钮电平（已去抖）。 *)
    b启动按钮 : BOOL;
    b暂停按钮 : BOOL;
    (* 上位机命令 2/3/4 已由 SEQ 去重，是独立的一扫描事件，
       不能与物理电平共用 R_TRIG，否则连续两帧命令会被合并。 *)
    b启动事件 : BOOL;
    b暂停事件 : BOOL;
    b恢复事件 : BOOL;
    b致命报警 : BOOL;
    b急停 : BOOL;
    b暂停报警 : BOOL;
    b预警 : BOOL;
    (* 由回收器回写：恢复进度与结果。 *)
    b暂停恢复中 : BOOL;
    b暂停恢复完成 : BOOL;
    b暂停恢复失败 : BOOL;
    b流程完成 : BOOL;
END_VAR
VAR_OUTPUT
    b运行指令 : BOOL;
    b期望运行 : BOOL;
    b暂停中 : BOOL;
    b自动模式 : BOOL;
    b手动模式 : BOOL;
    b自动可运行 : BOOL;
    (* 电平请求：置位启动暂停恢复，恢复完成后由本块清除。 *)
    b暂停恢复请求 : BOOL;
    b报警灯 : BOOL;
    b运行灯 : BOOL;
    b待机灯 : BOOL;
END_VAR
VAR
    rt启动 : R_TRIG;
    rt暂停 : R_TRIG;
END_VAR

rt启动(CLK := b启动按钮);
rt暂停(CLK := b暂停按钮);

b报警灯 := b致命报警 OR b暂停报警 OR b预警;
b自动可运行 := b初始化完成
    AND b系统复位完成
    AND NOT b系统复位中
    AND NOT b系统复位失败
    AND NOT b致命报警
    AND NOT b暂停恢复中
    AND NOT b暂停恢复失败;

(* 优先级：硬故障 > 流程完成 > 初始化/复位 > 暂停 > 启动。 *)
IF b致命报警 THEN
    b运行指令 := FALSE;
    b期望运行 := FALSE;
    b暂停中 := FALSE;
    b暂停恢复请求 := FALSE;
ELSIF b流程完成 THEN
    b运行指令 := FALSE;
    b期望运行 := FALSE;
    b暂停中 := FALSE;
    b暂停恢复请求 := FALSE;
ELSIF (NOT b初始化完成) OR (NOT b系统复位完成) THEN
    b运行指令 := FALSE;
    b期望运行 := FALSE;
    b暂停中 := FALSE;
    b暂停恢复请求 := FALSE;
ELSIF b系统复位中 OR b系统复位失败 THEN
    b运行指令 := FALSE;
    b期望运行 := FALSE;
    b暂停中 := FALSE;
    b暂停恢复请求 := FALSE;
ELSE
    (* 暂停恢复是一次性握手：请求 -> 恢复中 -> 完成/失败。
       恢复期间保持请求电平，完成或失败后立即撤销，不会重复触发。 *)
    IF b暂停恢复失败 THEN
        b暂停恢复请求 := FALSE;
        IF NOT b暂停恢复中 THEN b暂停中 := TRUE; END_IF;
    ELSIF b暂停恢复完成 AND b暂停恢复请求 AND NOT b暂停恢复中 THEN
        b暂停恢复请求 := FALSE;
        b暂停中 := FALSE;
        b运行指令 := TRUE;
        b期望运行 := TRUE;
    END_IF;

    IF NOT b暂停恢复请求 AND NOT b暂停恢复中 THEN
        IF rt暂停.Q OR b暂停事件 THEN
            IF b运行指令 THEN
                b运行指令 := FALSE;
                b暂停中 := TRUE;
            END_IF;
        (* 同一扫描启动和暂停同时出现时，暂停优先。
           暂停中不接受启动：暂停必须经命令 4 的受控恢复退出，
           否则会绕过暂停快照回位直接重新运行。 *)
        ELSIF (rt启动.Q OR b启动事件)
        AND NOT b暂停中
        AND b自动可运行
        AND NOT b暂停报警 THEN
            b期望运行 := TRUE;
            b运行指令 := TRUE;
            b暂停中 := FALSE;
        (* 命令 4：暂停中的受控恢复请求。 *)
        ELSIF b恢复事件 AND b暂停中 AND b自动可运行 AND NOT b暂停报警 THEN
            b暂停恢复请求 := TRUE;
        END_IF;
    END_IF;

    (* 急停在任何恢复阶段都立即撤销请求；恢复结果由回收器置失败。 *)
    IF b急停 THEN b暂停恢复请求 := FALSE; END_IF;
END_IF;

(* 模式只描述当前控制归属，不代表动作已经获得安全许可。 *)
b自动模式 := b运行指令;
b手动模式 := NOT b运行指令 AND NOT b急停;
b运行灯 := b运行指令;
b待机灯 := NOT b运行指令 AND NOT b报警灯;
END_FUNCTION_BLOCK
